// TIA Portal V21 export
// export: Created 2026-11-11T00:48:14.6140209Z, ExportSetting WithDefaults, DisplayName Totally Integrated Automation Portal, DisplayVersion V21 Update 3, DisplayName STEP 7 Professional, DisplayVersion V21 Update 3, DisplayName STEP 7 Safety, DisplayVersion V21, DisplayName Tech WebApplication, DisplayVersion V21, DisplayName WinCC Basic/Comfort/Advanced, DisplayVersion V21 Update 3, DisplayName WinCC Unified, DisplayVersion V21 Update 3
FUNCTION_BLOCK "FB_Scl_sl034"   // FB56, SCL
{ S7_Optimized_Access := 'TRUE' }
VERSION : 0.1
// stored: AutoNumber true, IsIECCheckEnabled false, IsRetainMemResEnabled false, MemoryReserve 100, SetENOAutomatically false, UDAEnableTagReadback false
   VAR_INPUT
      v_in : Real;
   END_VAR
   VAR_OUTPUT
      v_ret : Real;
   END_VAR
BEGIN
   #v_ret := TAN(IN := #v_in);
END_FUNCTION_BLOCK
